Fanuc KAREL source: KT00990.KL

PROGRAM KT00990
%NOLOCKGROUP
VAR
  H1: ARRAY[2] OF SHORT
  H2: ARRAY[2] OF SHORT
  CFG: CONFIG
  OUT: XYZWPREXT
BEGIN
  H1[1] = 2
  H2[1] = 3
  H1[1] = 2
  H2[1] = 3
  CFG.CFG_FLIP = TRUE
  OUT = POS(H1[1], H1[1], H1[1], H1[1], H1[1], H1[1], CFG)
END KT00990
